(* IEC 61131-3 sources: llm-plc-st-eval/data/processed_v2_primera/claude-sonnet-4-6/B5/zero_shot, 3 files *)

(* ---- ejec_1.st ---- *)
FUNCTION_BLOCK FB_Ventilador
VAR_INPUT
    quemadorOn : BOOL; (* Señal del quemador: TRUE = encendido *)
END_VAR

VAR_OUTPUT
    ventilador : BOOL; (* Salida del ventilador: TRUE = funcionando *)
END_VAR

VAR
    tPostEnfriamiento : TON;  (* Temporizador de post-enfriamiento *)
END_VAR

(*
    Lógica:
    - Si el quemador está encendido, el ventilador funciona y el temporizador se mantiene reseteado.
    - Al apagarse el quemador, el temporizador inicia y el ventilador sigue funcionando.
    - Transcurridos 30 s, el temporizador expira y el ventilador se detiene.
*)

(* Activar temporizador solo cuando el quemador está apagado *)
tPostEnfriamiento(
    IN  := NOT quemadorOn,
    PT  := T#30S
);

(* El ventilador funciona si el quemador está ON o si el temporizador aún no expiró *)
ventilador := quemadorOn OR NOT tPostEnfriamiento.Q;

(* ---- ejec_2.st ---- *)
FUNCTION_BLOCK FB_Ventilador
VAR_INPUT
    quemadorOn : BOOL; (* Señal del quemador: TRUE = encendido *)
END_VAR

VAR_OUTPUT
    ventilador : BOOL; (* Salida del ventilador: TRUE = funcionando *)
END_VAR

VAR
    tonPostApagado : TON;  (* Temporizador de retardo al apagado *)
END_VAR

(*
    Lógica:
    - Si el quemador está encendido, el ventilador funciona y el temporizador se mantiene reseteado.
    - Al apagarse el quemador, el temporizador comienza a contar 30 segundos.
    - Mientras el temporizador no haya expirado, el ventilador sigue funcionando.
    - Una vez transcurridos los 30 segundos, el ventilador se detiene.
*)

(* Activar temporizador solo cuando el quemador está apagado *)
tonPostApagado(
    IN  := NOT quemadorOn,
    PT  := T#30S
);

(* El ventilador funciona si el quemador está ON o si el temporizador aún no ha expirado *)
ventilador := quemadorOn OR NOT tonPostApagado.Q;

END_FUNCTION_BLOCK

(* ---- ejec_3.st ---- *)
FUNCTION_BLOCK FB_Ventilador
VAR_INPUT
    quemadorOn : BOOL; (* Señal del quemador: TRUE = encendido *)
END_VAR

VAR_OUTPUT
    ventilador : BOOL; (* Salida del ventilador: TRUE = funcionando *)
END_VAR

VAR
    tonPostApagado : TON;  (* Temporizador de retardo al apagado *)
END_VAR

(*
    Lógica:
    - Si el quemador está encendido, el ventilador funciona y el temporizador se mantiene reseteado.
    - Al apagarse el quemador, el temporizador comienza a contar 30 segundos.
    - Cuando el temporizador completa los 30 segundos (Q = TRUE), el ventilador se detiene.
*)

(* Activar temporizador solo cuando el quemador está apagado *)
tonPostApagado(
    IN  := NOT quemadorOn,
    PT  := T#30S
);

(* El ventilador funciona si el quemador está encendido
   O si el temporizador aún no ha completado los 30 segundos *)
ventilador := quemadorOn OR NOT tonPostApagado.Q;

END_FUNCTION_BLOCK
